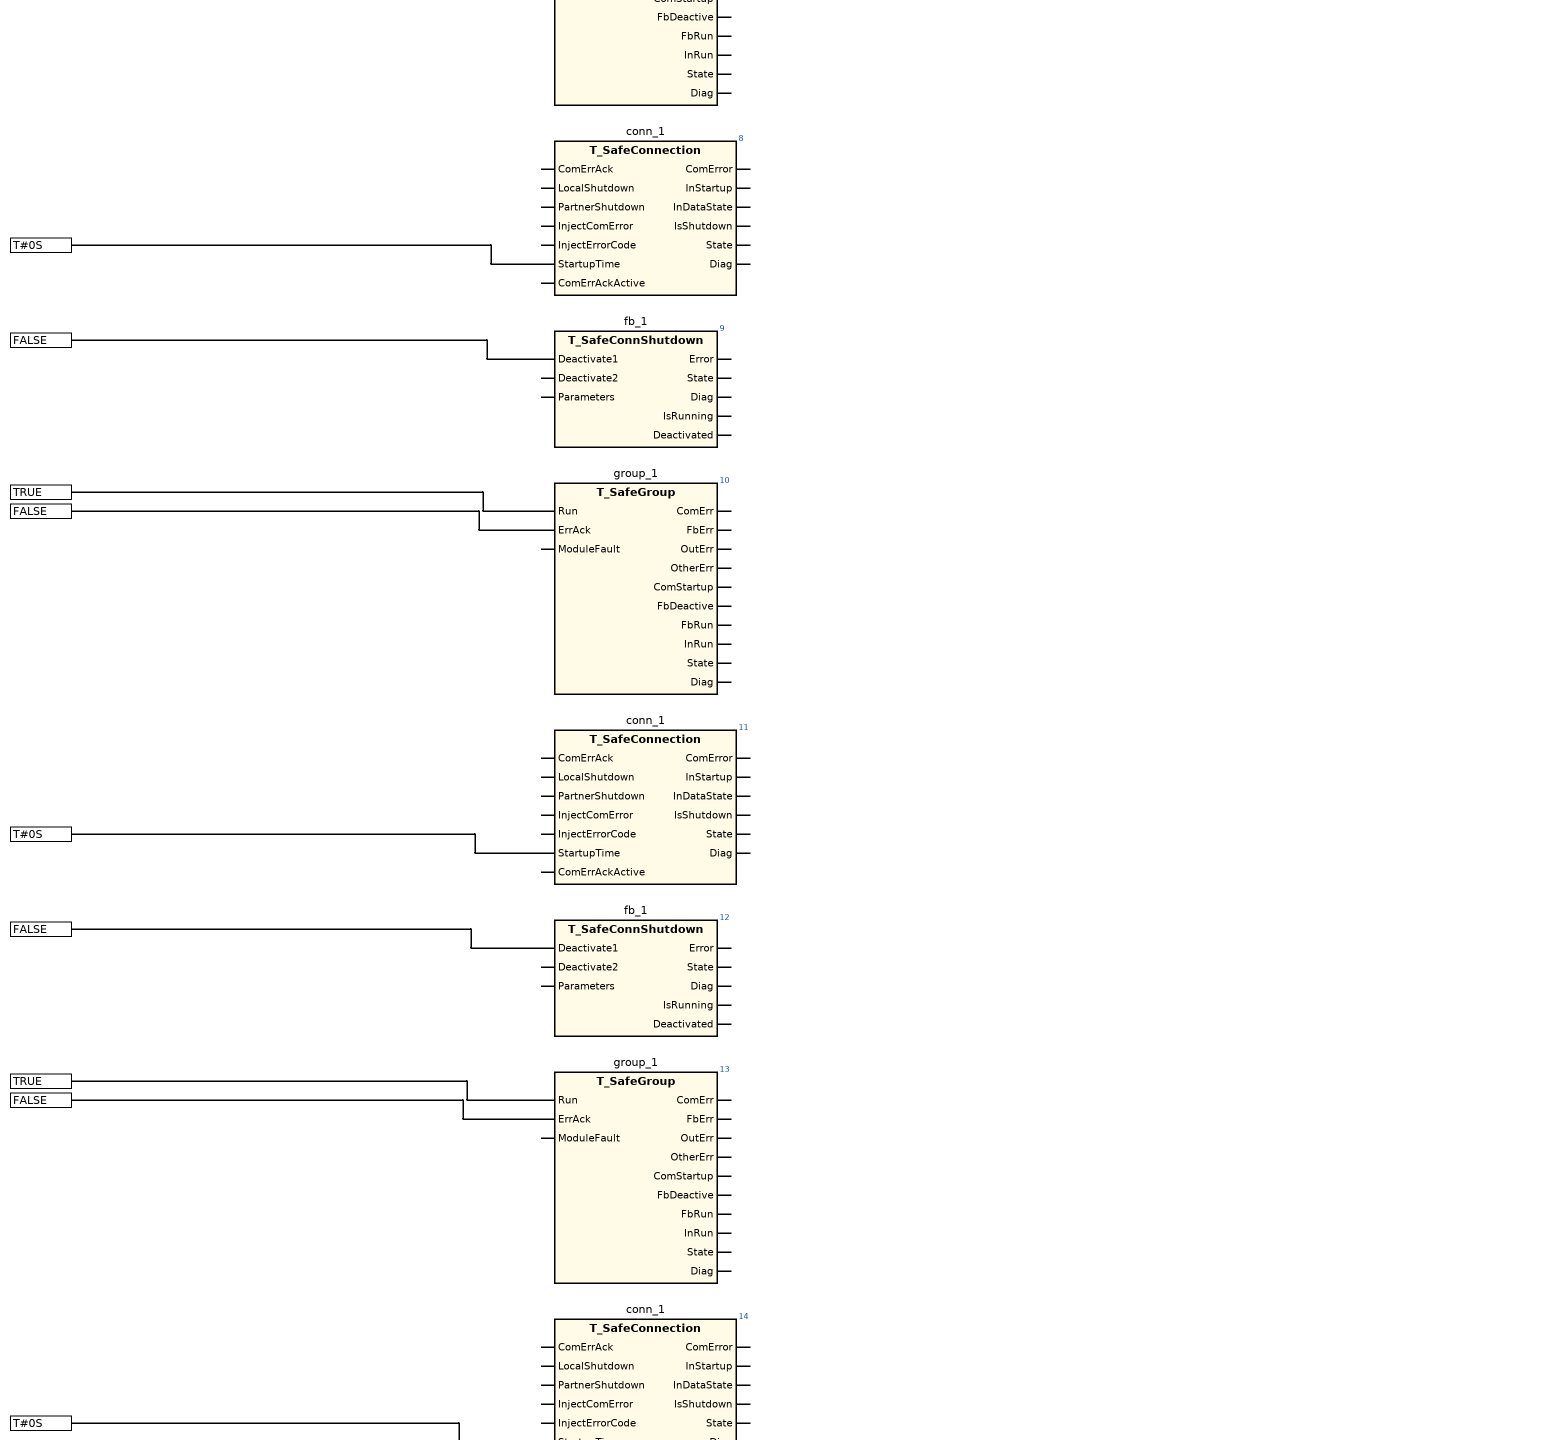
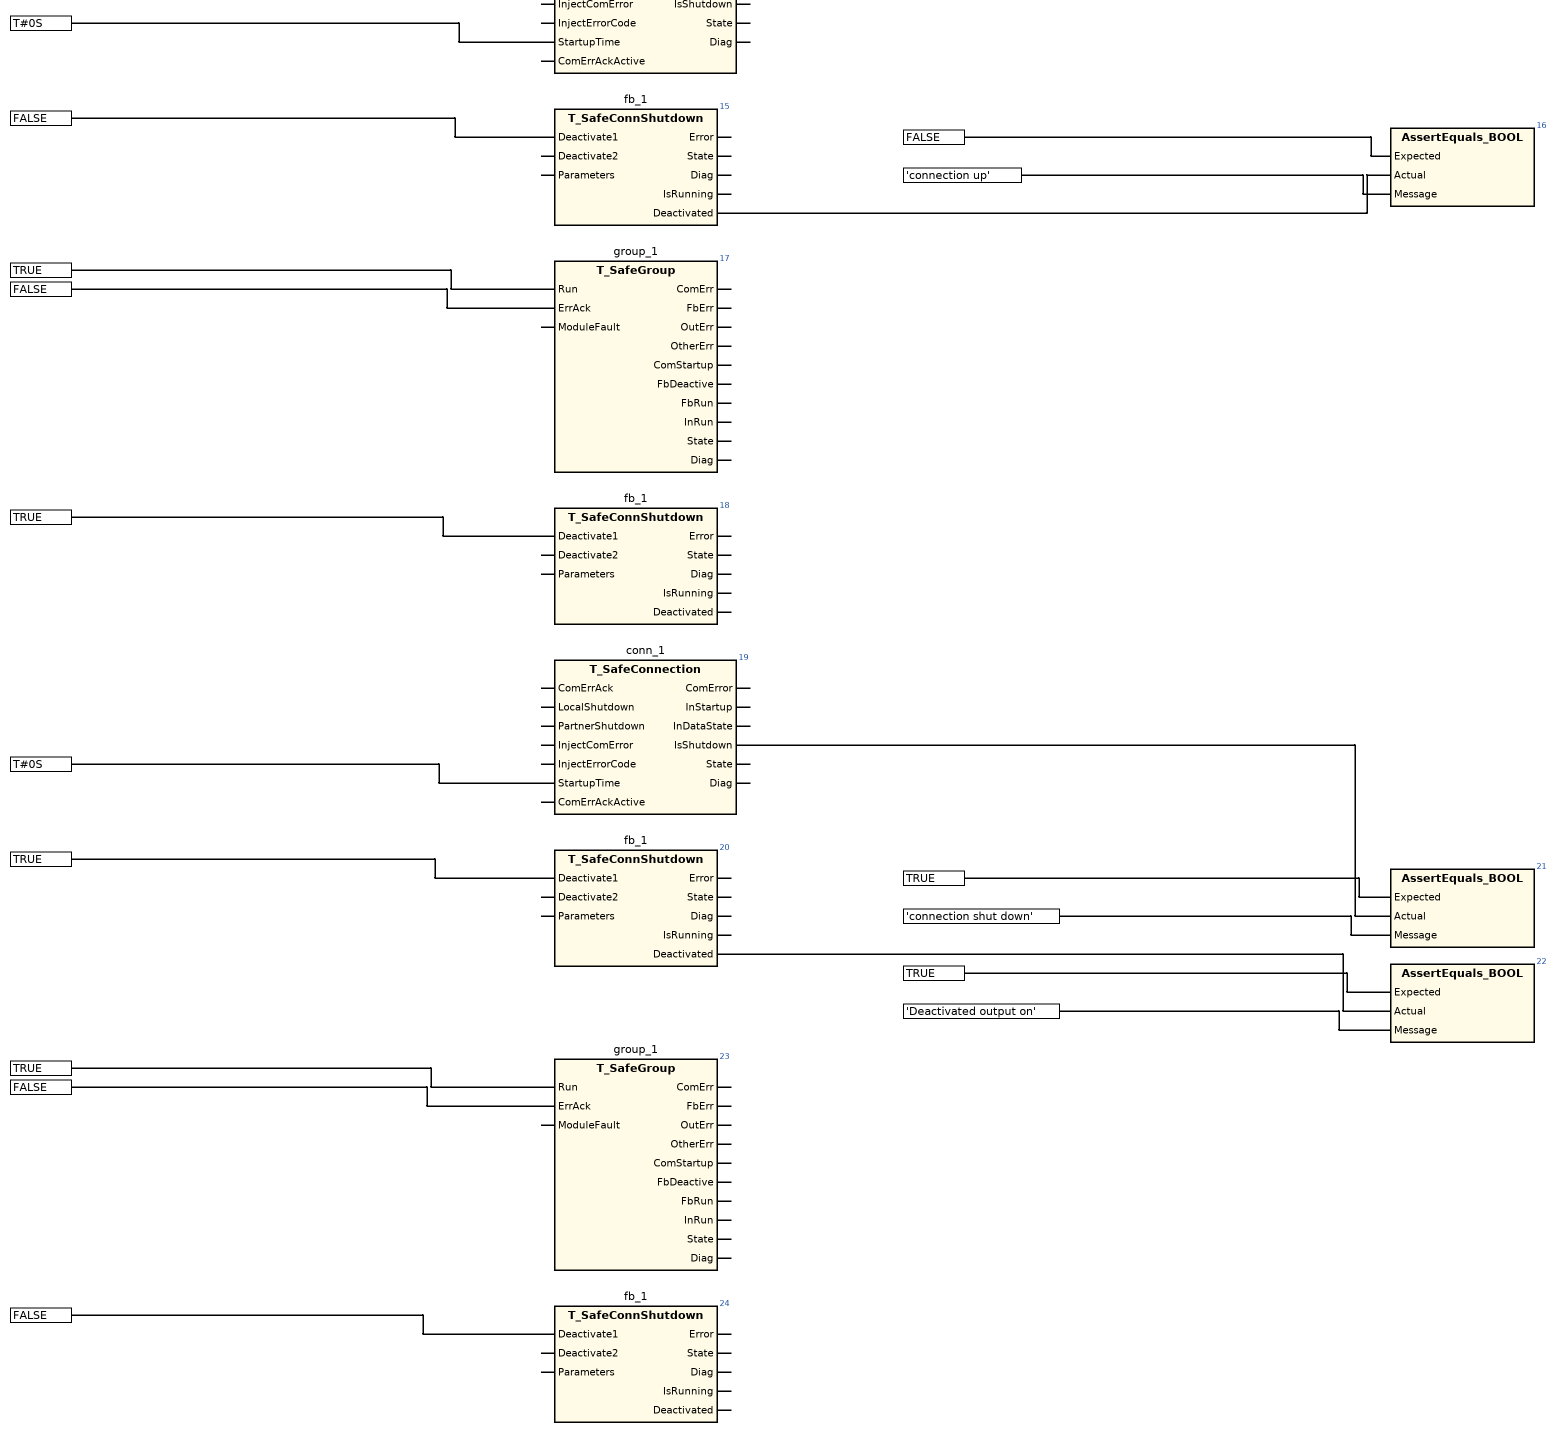
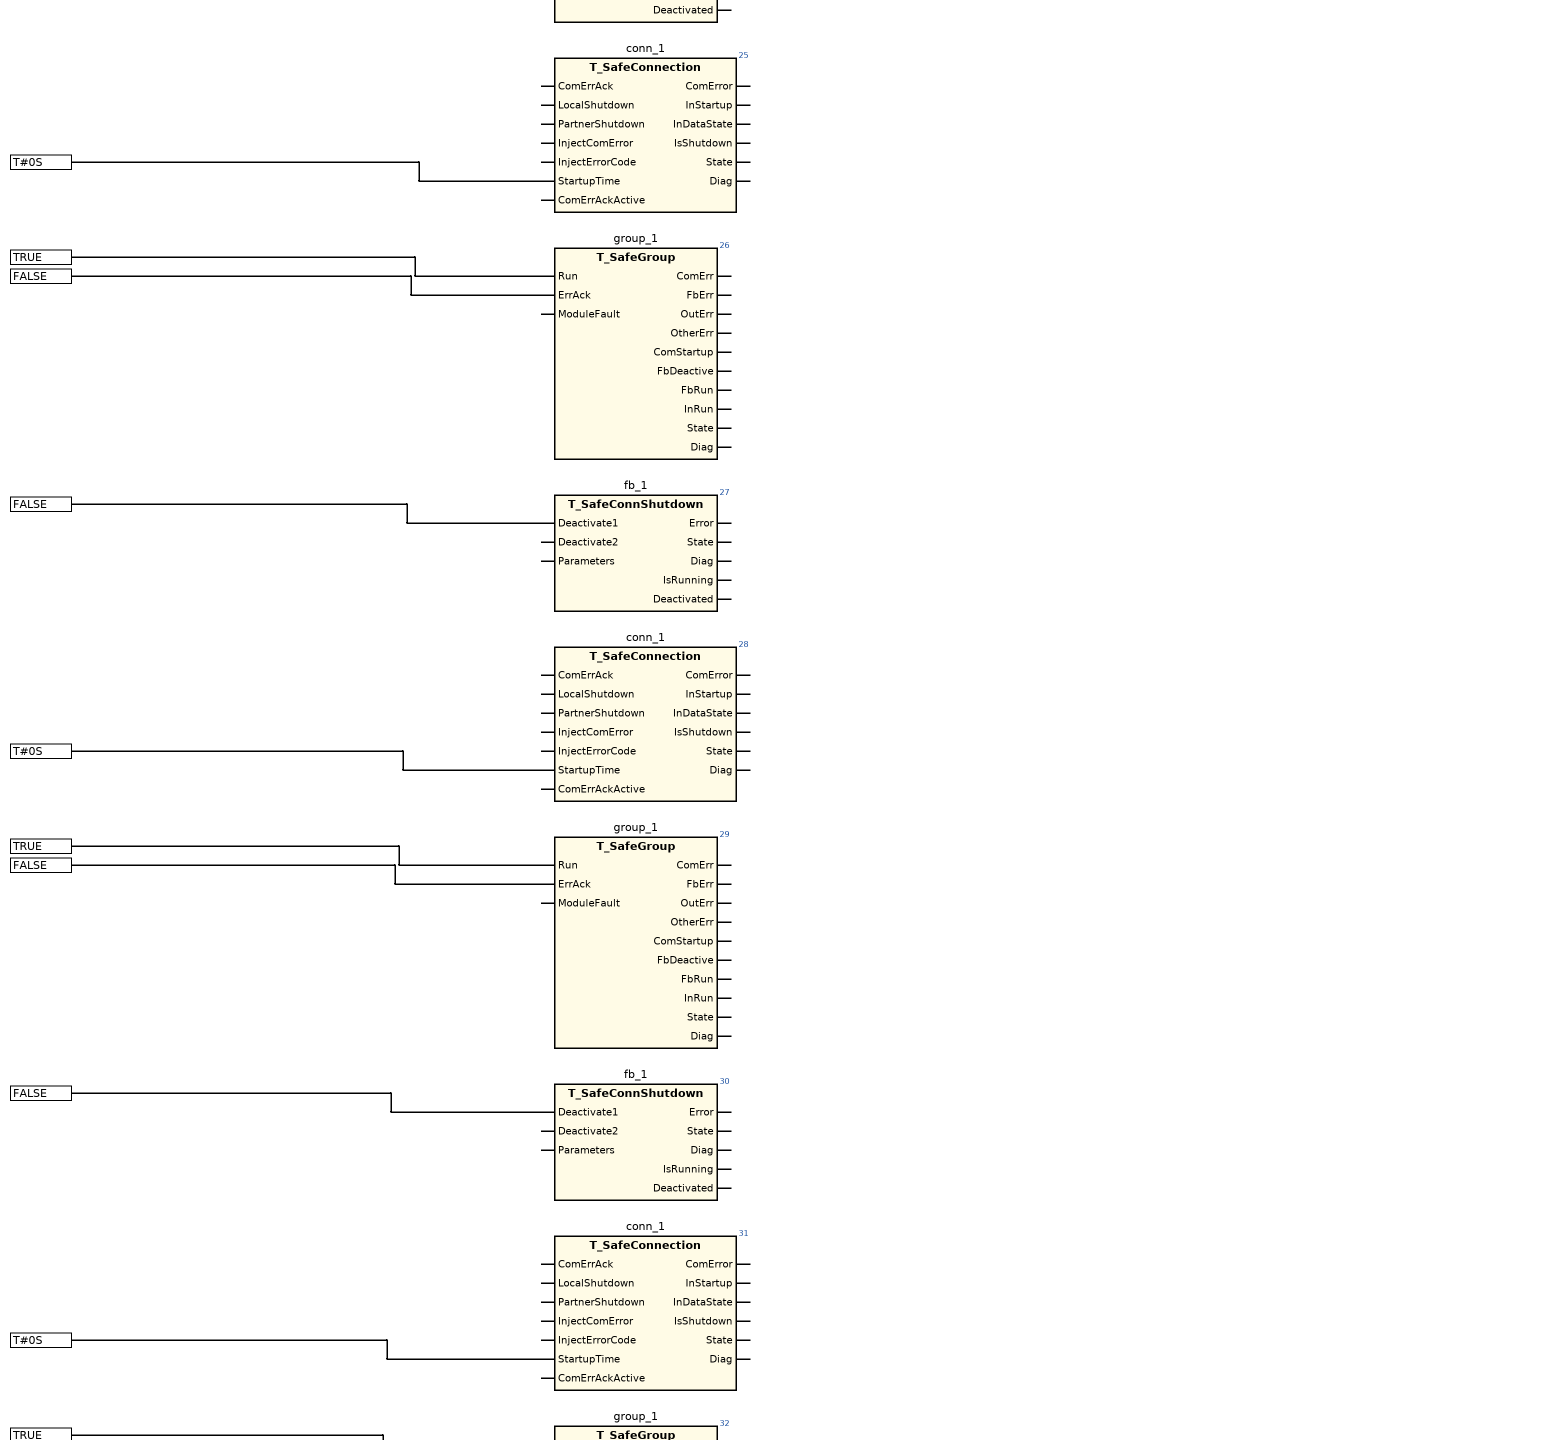
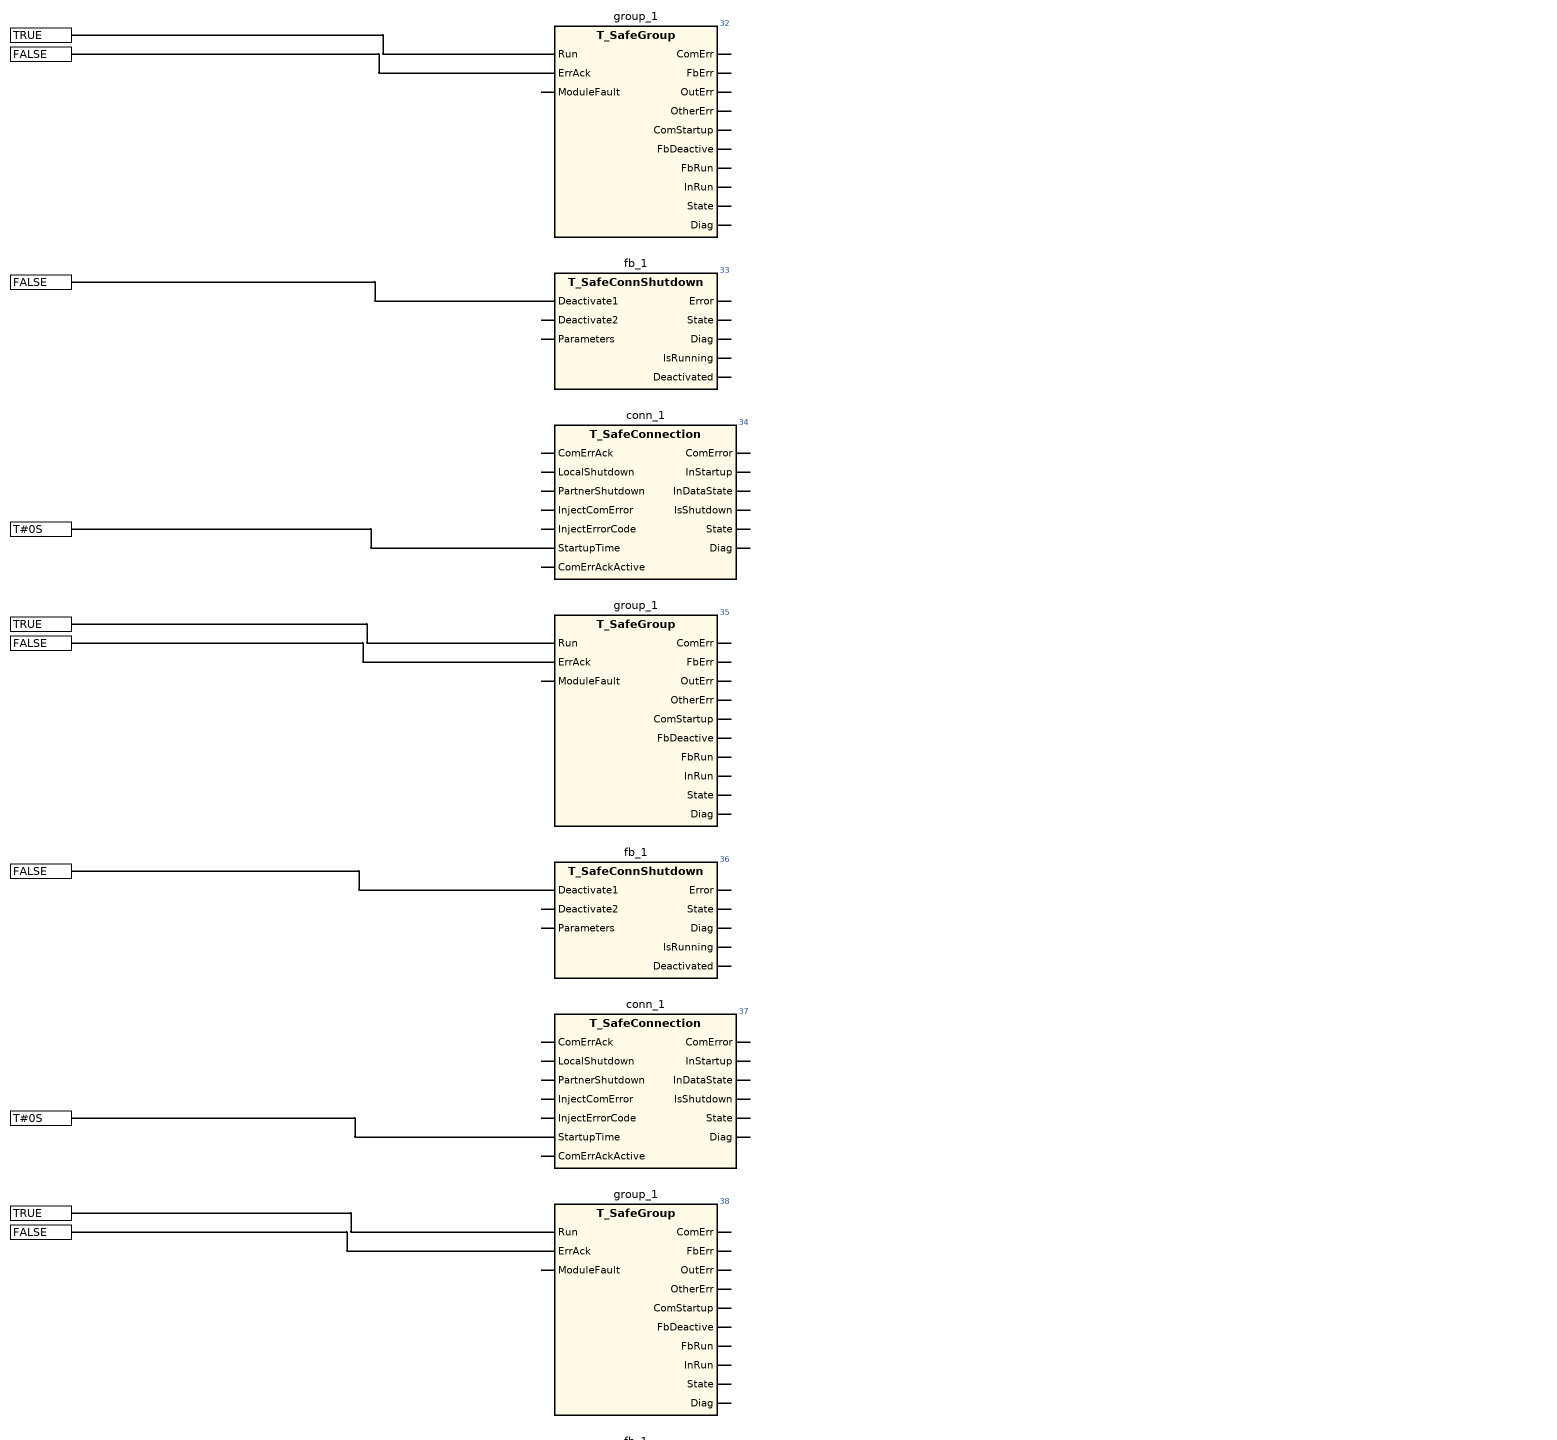
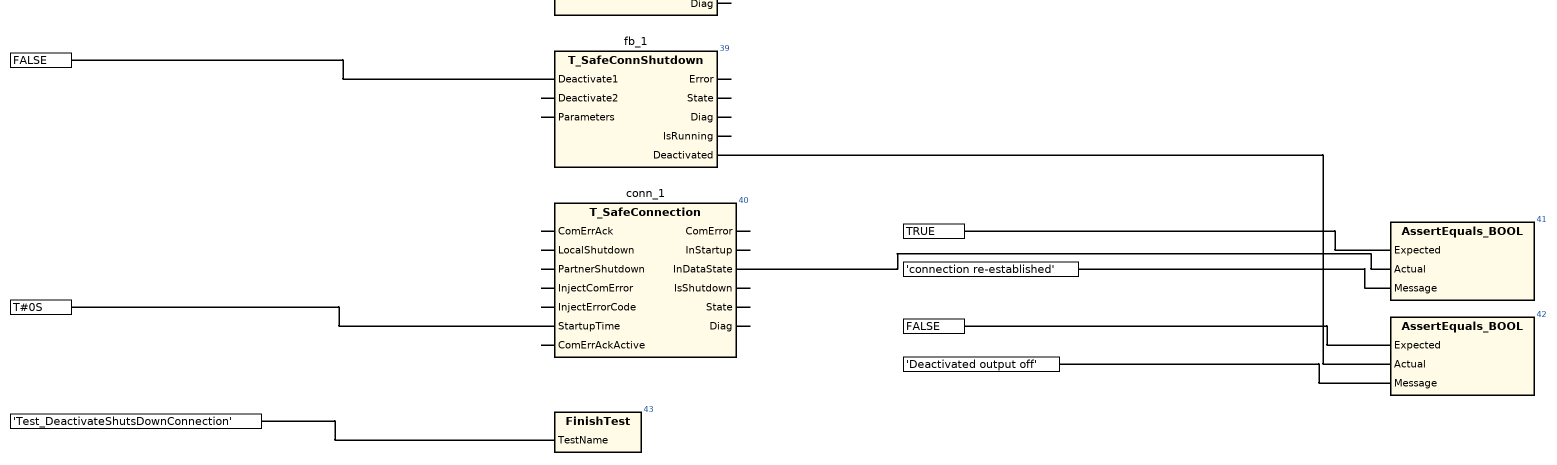
StartTest(TestName := 'Test_DeactivateShutsDownConnection');
group_1(Run := TRUE, ErrAck := FALSE); // T_SafeGroup
conn_1(StartupTime := T#0S); // T_SafeConnection
fb_1(Deactivate1 := FALSE); // T_SafeConnShutdown
group_1(Run := TRUE, ErrAck := FALSE); // T_SafeGroup
conn_1(StartupTime := T#0S); // T_SafeConnection
fb_1(Deactivate1 := FALSE); // T_SafeConnShutdown
group_1(Run := TRUE, ErrAck := FALSE); // T_SafeGroup
conn_1(StartupTime := T#0S); // T_SafeConnection
fb_1(Deactivate1 := FALSE); // T_SafeConnShutdown
group_1(Run := TRUE, ErrAck := FALSE); // T_SafeGroup
conn_1(StartupTime := T#0S); // T_SafeConnection
fb_1(Deactivate1 := FALSE); // T_SafeConnShutdown
group_1(Run := TRUE, ErrAck := FALSE); // T_SafeGroup
conn_1(StartupTime := T#0S); // T_SafeConnection
fb_1(Deactivate1 := FALSE); // T_SafeConnShutdown
AssertEquals_BOOL(Expected := FALSE, Actual := fb_1.Deactivated, Message := 'connection up');
group_1(Run := TRUE, ErrAck := FALSE); // T_SafeGroup
fb_1(Deactivate1 := TRUE); // T_SafeConnShutdown
conn_1(StartupTime := T#0S); // T_SafeConnection
fb_1(Deactivate1 := TRUE); // T_SafeConnShutdown
AssertEquals_BOOL(Expected := TRUE, Actual := conn_1.IsShutdown, Message := 'connection shut down');
AssertEquals_BOOL(Expected := TRUE, Actual := fb_1.Deactivated, Message := 'Deactivated output on');
group_1(Run := TRUE, ErrAck := FALSE); // T_SafeGroup
fb_1(Deactivate1 := FALSE); // T_SafeConnShutdown
conn_1(StartupTime := T#0S); // T_SafeConnection
group_1(Run := TRUE, ErrAck := FALSE); // T_SafeGroup
fb_1(Deactivate1 := FALSE); // T_SafeConnShutdown
conn_1(StartupTime := T#0S); // T_SafeConnection
group_1(Run := TRUE, ErrAck := FALSE); // T_SafeGroup
fb_1(Deactivate1 := FALSE); // T_SafeConnShutdown
conn_1(StartupTime := T#0S); // T_SafeConnection
group_1(Run := TRUE, ErrAck := FALSE); // T_SafeGroup
fb_1(Deactivate1 := FALSE); // T_SafeConnShutdown
conn_1(StartupTime := T#0S); // T_SafeConnection
group_1(Run := TRUE, ErrAck := FALSE); // T_SafeGroup
fb_1(Deactivate1 := FALSE); // T_SafeConnShutdown
conn_1(StartupTime := T#0S); // T_SafeConnection
group_1(Run := TRUE, ErrAck := FALSE); // T_SafeGroup
fb_1(Deactivate1 := FALSE); // T_SafeConnShutdown
conn_1(StartupTime := T#0S); // T_SafeConnection
AssertEquals_BOOL(Expected := TRUE, Actual := conn_1.InDataState, Message := 'connection re-established');
AssertEquals_BOOL(Expected := FALSE, Actual := fb_1.Deactivated, Message := 'Deactivated output off');
FinishTest(TestName := 'Test_DeactivateShutsDownConnection');
END_METHOD

END_FUNCTION_BLOCK

// Tests/T_SafeGroup_Tests_CFC
    // CFC twin of T_SafeGroup_Tests: the same tests drawn as CFC diagrams, the way a TwinSAFE project is authored.
    FUNCTION_BLOCK T_SafeGroup_Tests_CFC EXTENDS T_SafeCfcTestSuite
    VAR
    // Test_StopWhenRunFalse
    group_1 : T_SafeGroup;
    fb_1 : T_SafeAnd(group := group_1);
    // Test_RunsFunctionBlocksWithoutConnections
    group_2 : T_SafeGroup;
    fb_2 : T_SafeAnd(group := group_2);
    // Test_FbErrorStopsGroupAndErrAckRecovers
    group_3 : T_SafeGroup;
    eStop_3 : T_SafeEStop(group := group_3);
    andFb_3 : T_SafeAnd(group := group_3);
    // Test_ConnectionStartupAndComError
    group_4 : T_SafeGroup;
    terminal_4 : T_SafeInputTerminal(group := group_4);
    t1a_4 : TON;
    t1b_4 : TON;
    t2b_4 : TON;
    trig1a_4 : R_TRIG;
    trig1b_4 : R_TRIG;
    trig2b_4 : R_TRIG;
    t3_4 : TON;
    trig3_4 : R_TRIG;
    t0_4 : TON;
    t1_4 : TON;
    t2_4 : TON;
    t4_4 : TON;
    trig0_4 : R_TRIG;
    trig1_4 : R_TRIG;
    trig2_4 : R_TRIG;
    trig4_4 : R_TRIG;
END_VAR

Test_StopWhenRunFalse();
Test_RunsFunctionBlocksWithoutConnections();
Test_FbErrorStopsGroupAndErrAckRecovers();
Test_ConnectionStartupAndComError();

METHOD PRIVATE Test_ConnectionStartupAndComError
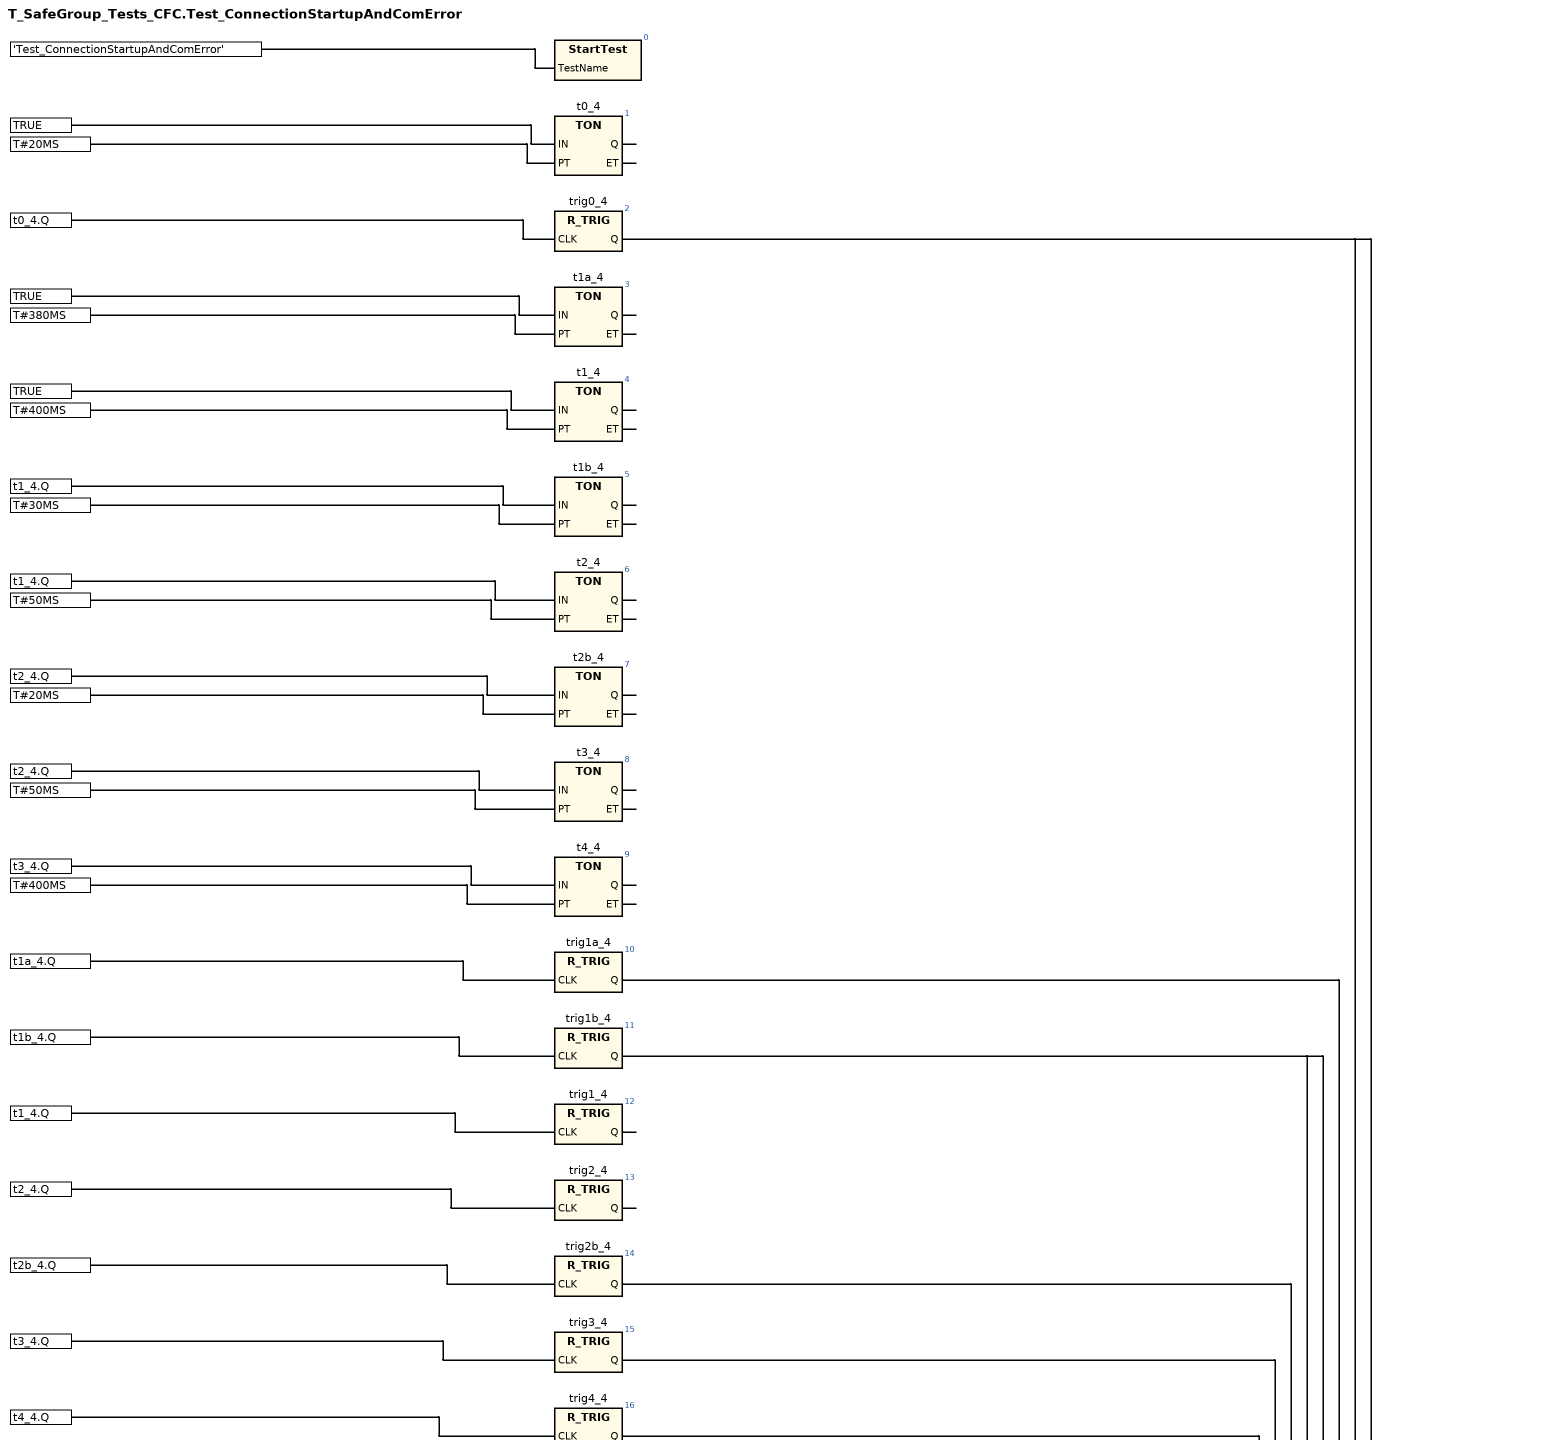
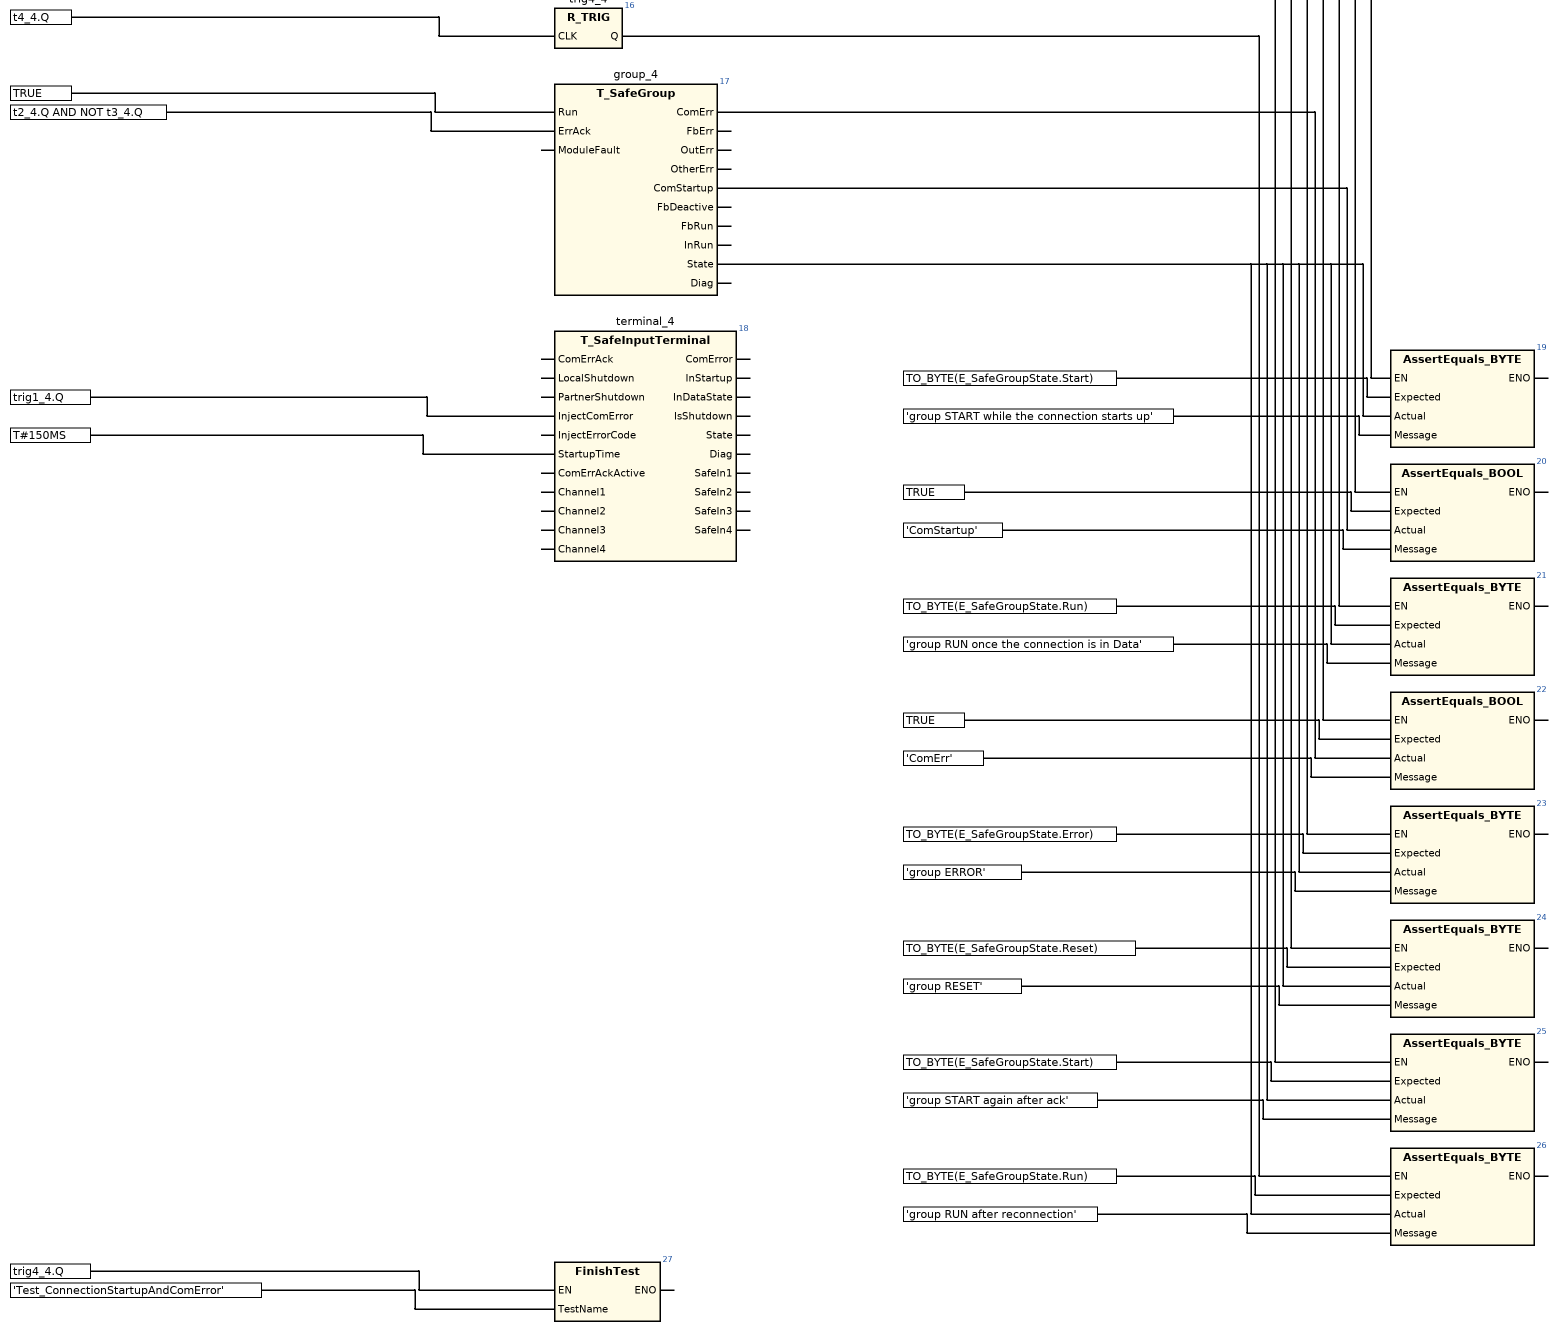
StartTest(TestName := 'Test_ConnectionStartupAndComError');
t0_4(IN := TRUE, PT := T#20MS); // TON
trig0_4(CLK := t0_4.Q); // R_TRIG
t1a_4(IN := TRUE, PT := T#380MS); // TON
t1_4(IN := TRUE, PT := T#400MS); // TON
t1b_4(IN := t1_4.Q, PT := T#30MS); // TON
t2_4(IN := t1_4.Q, PT := T#50MS); // TON
t2b_4(IN := t2_4.Q, PT := T#20MS); // TON
t3_4(IN := t2_4.Q, PT := T#50MS); // TON
t4_4(IN := t3_4.Q, PT := T#400MS); // TON
trig1a_4(CLK := t1a_4.Q); // R_TRIG
trig1b_4(CLK := t1b_4.Q); // R_TRIG
trig1_4(CLK := t1_4.Q); // R_TRIG
trig2_4(CLK := t2_4.Q); // R_TRIG
trig2b_4(CLK := t2b_4.Q); // R_TRIG
trig3_4(CLK := t3_4.Q); // R_TRIG
trig4_4(CLK := t4_4.Q); // R_TRIG
group_4(Run := TRUE, ErrAck := t2_4.Q AND NOT t3_4.Q); // T_SafeGroup
terminal_4(InjectComError := trig1_4.Q, StartupTime := T#150MS); // T_SafeInputTerminal
IF trig0_4.Q THEN AssertEquals_BYTE(Expected := TO_BYTE(E_SafeGroupState.Start), Actual := group_4.State, Message := 'group START while the connection starts up'); END_IF
IF trig0_4.Q THEN AssertEquals_BOOL(Expected := TRUE, Actual := group_4.ComStartup, Message := 'ComStartup'); END_IF
IF trig1a_4.Q THEN AssertEquals_BYTE(Expected := TO_BYTE(E_SafeGroupState.Run), Actual := group_4.State, Message := 'group RUN once the connection is in Data'); END_IF
IF trig1b_4.Q THEN AssertEquals_BOOL(Expected := TRUE, Actual := group_4.ComErr, Message := 'ComErr'); END_IF
IF trig1b_4.Q THEN AssertEquals_BYTE(Expected := TO_BYTE(E_SafeGroupState.Error), Actual := group_4.State, Message := 'group ERROR'); END_IF
IF trig2b_4.Q THEN AssertEquals_BYTE(Expected := TO_BYTE(E_SafeGroupState.Reset), Actual := group_4.State, Message := 'group RESET'); END_IF
IF trig3_4.Q THEN AssertEquals_BYTE(Expected := TO_BYTE(E_SafeGroupState.Start), Actual := group_4.State, Message := 'group START again after ack'); END_IF
IF trig4_4.Q THEN AssertEquals_BYTE(Expected := TO_BYTE(E_SafeGroupState.Run), Actual := group_4.State, Message := 'group RUN after reconnection'); END_IF
IF trig4_4.Q THEN FinishTest(TestName := 'Test_ConnectionStartupAndComError'); END_IF
END_METHOD

METHOD PRIVATE Test_FbErrorStopsGroupAndErrAckRecovers
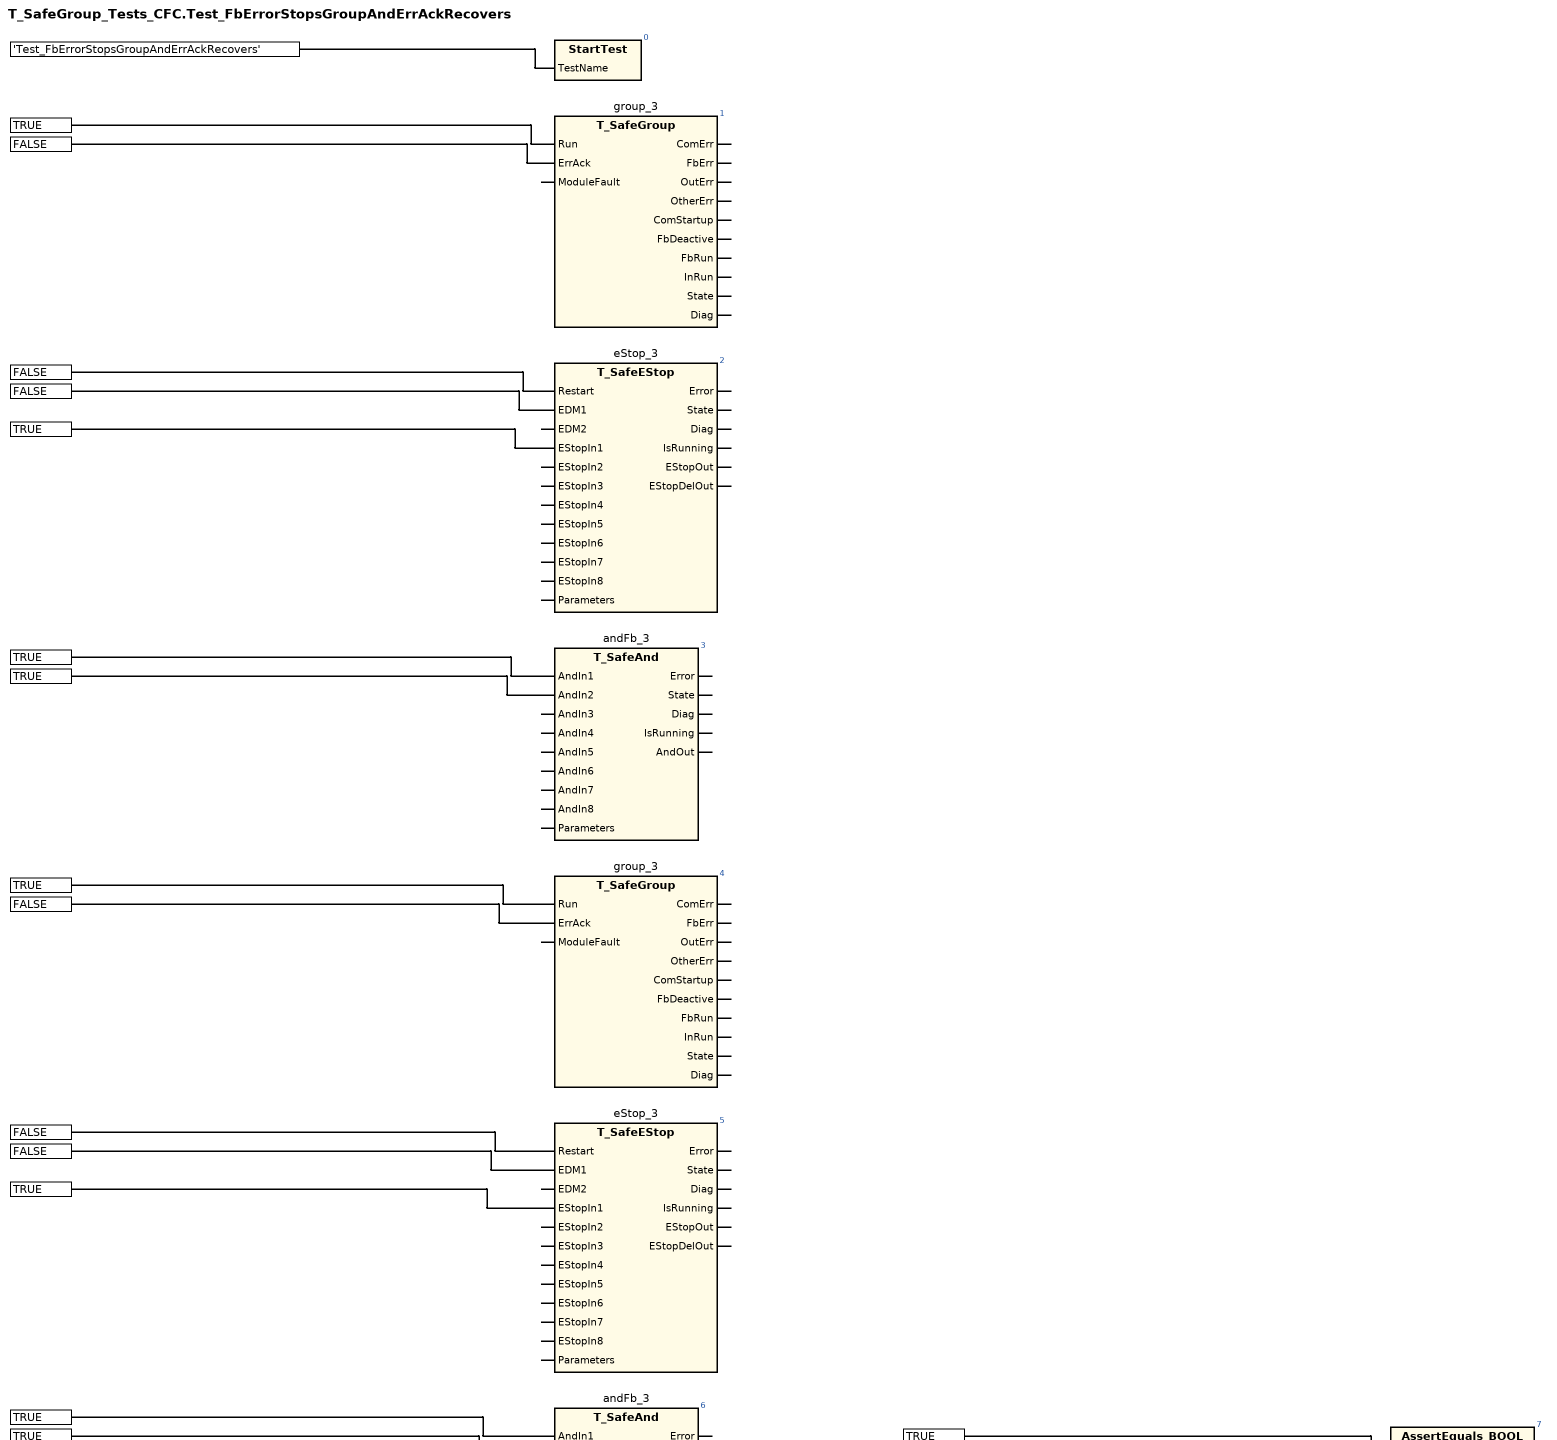
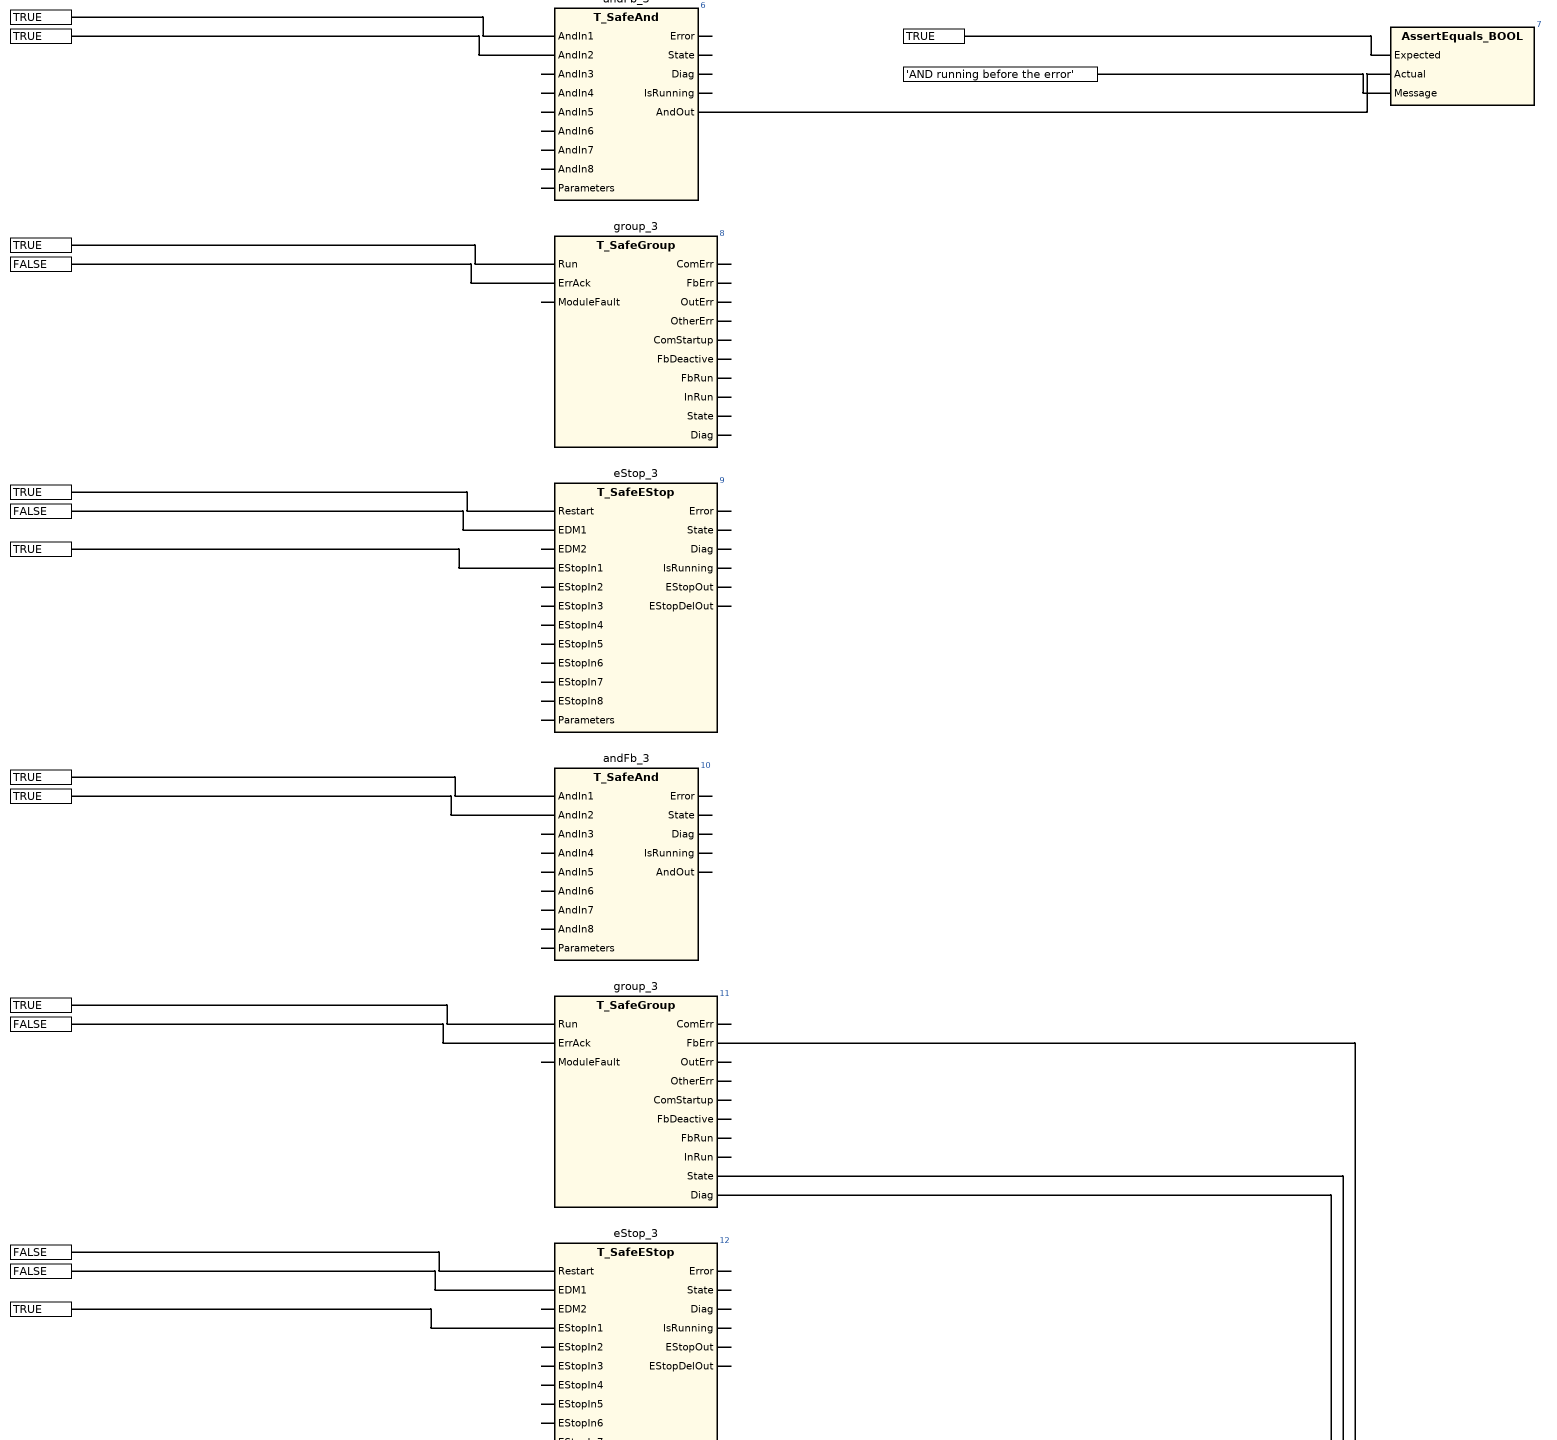
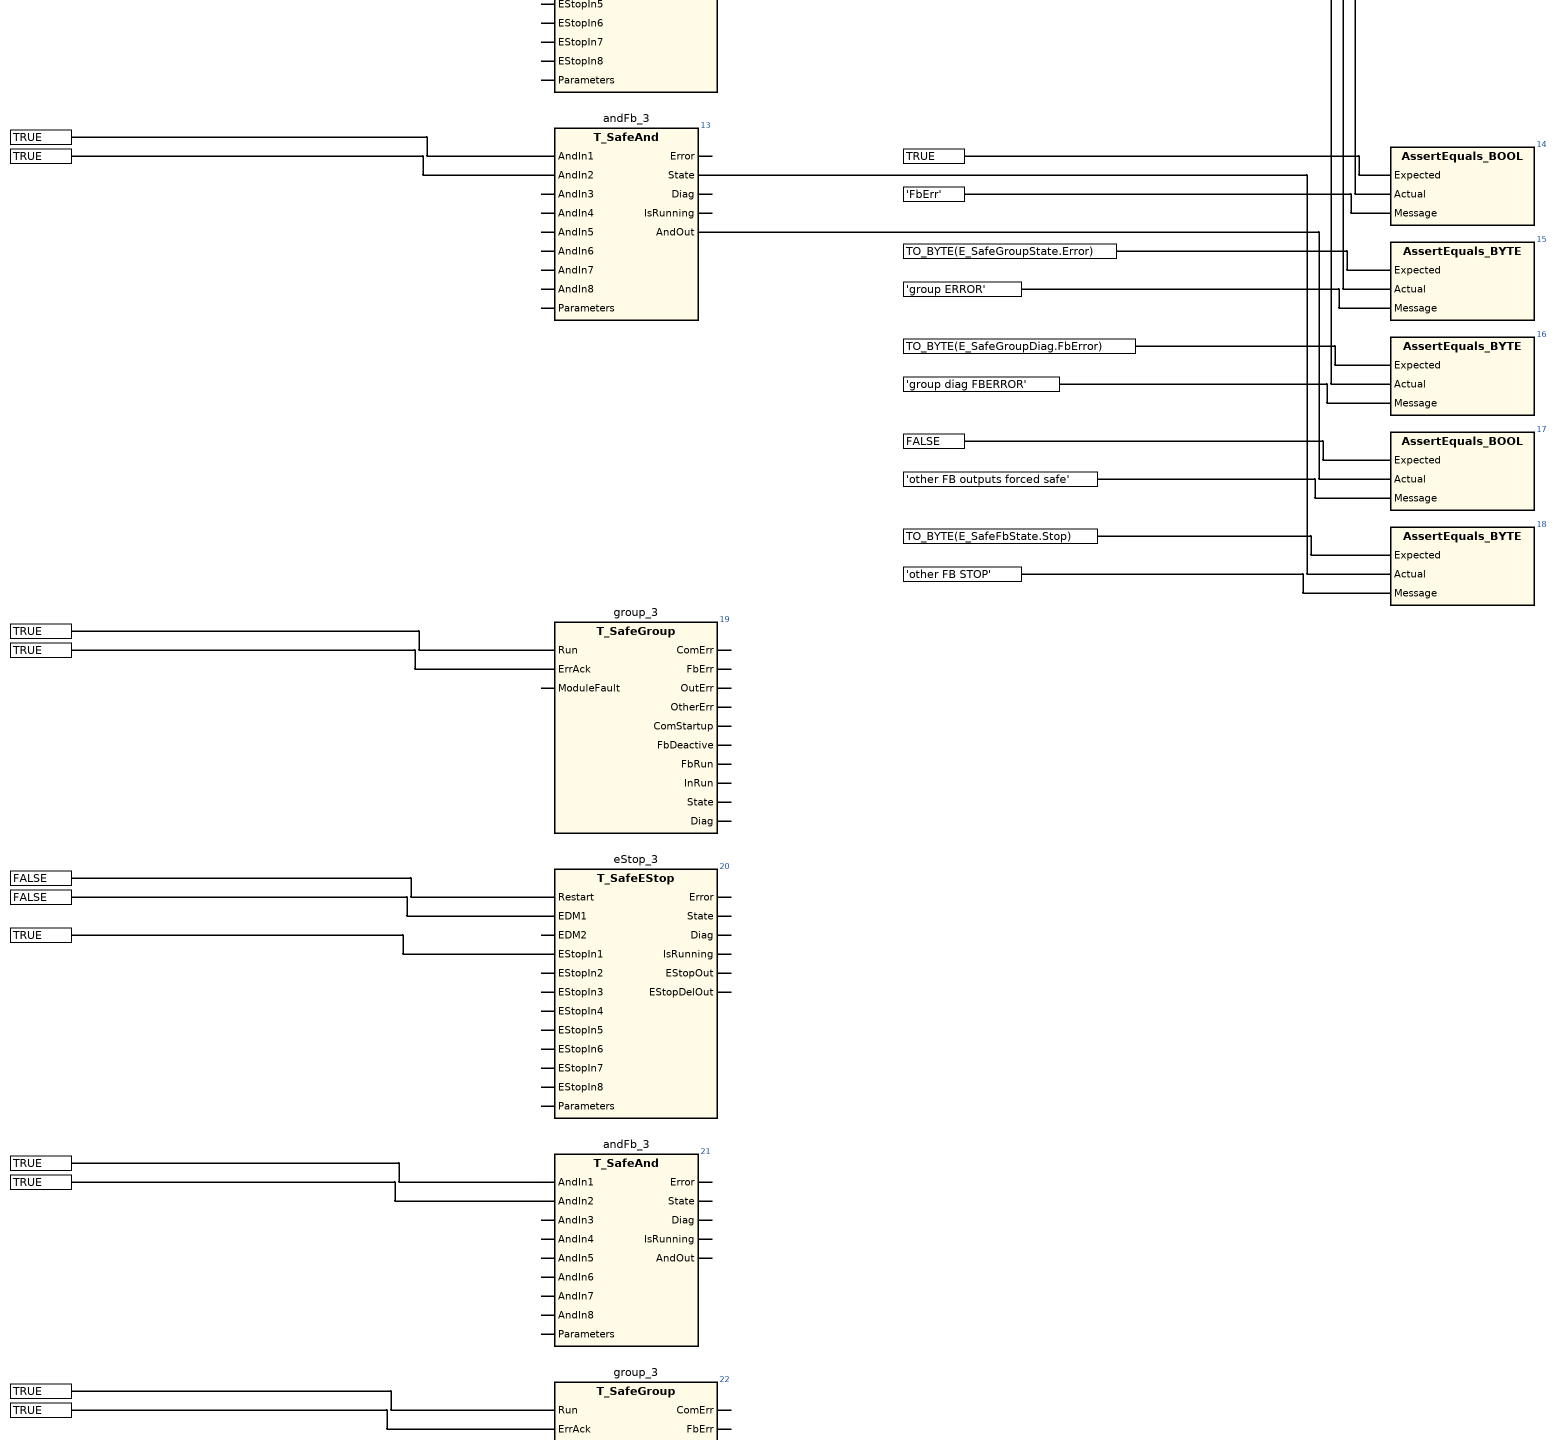
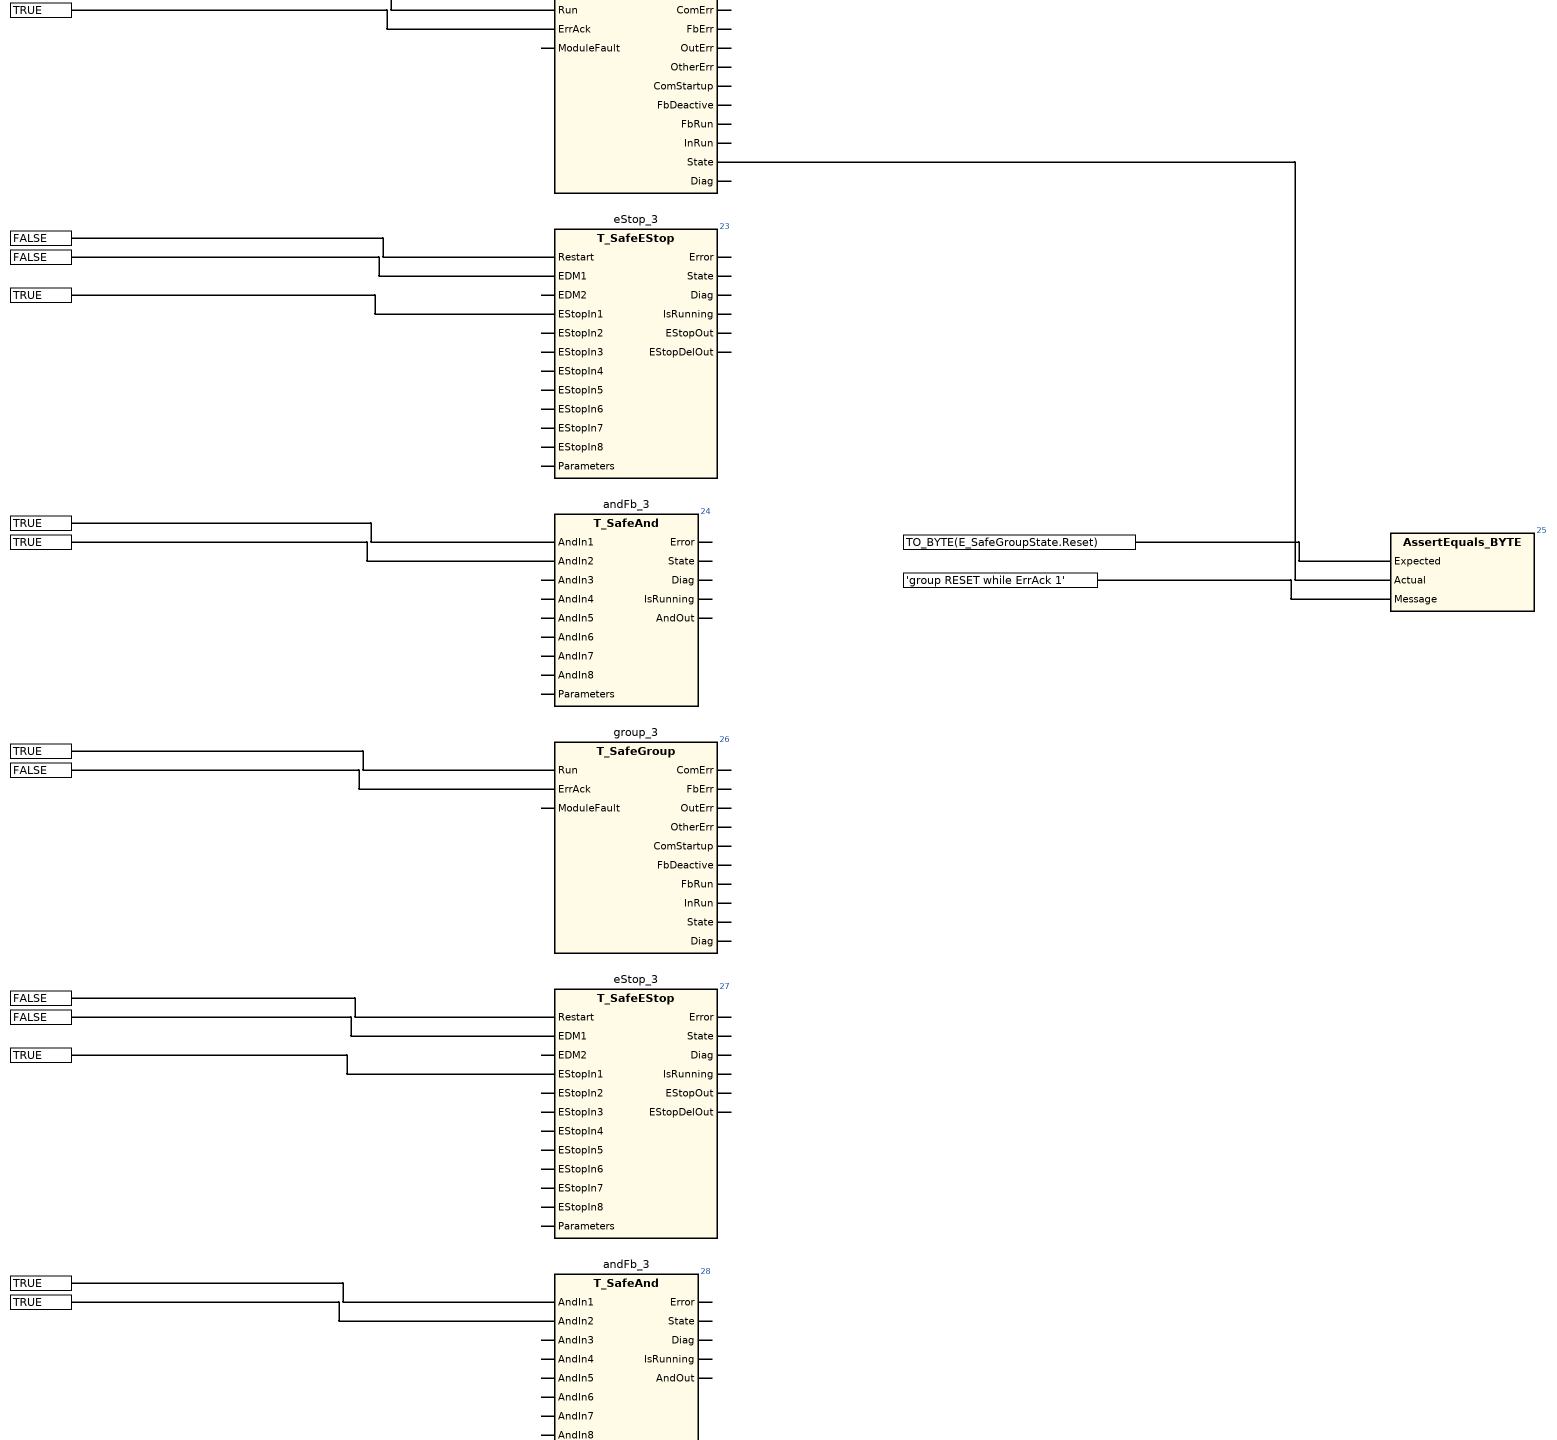
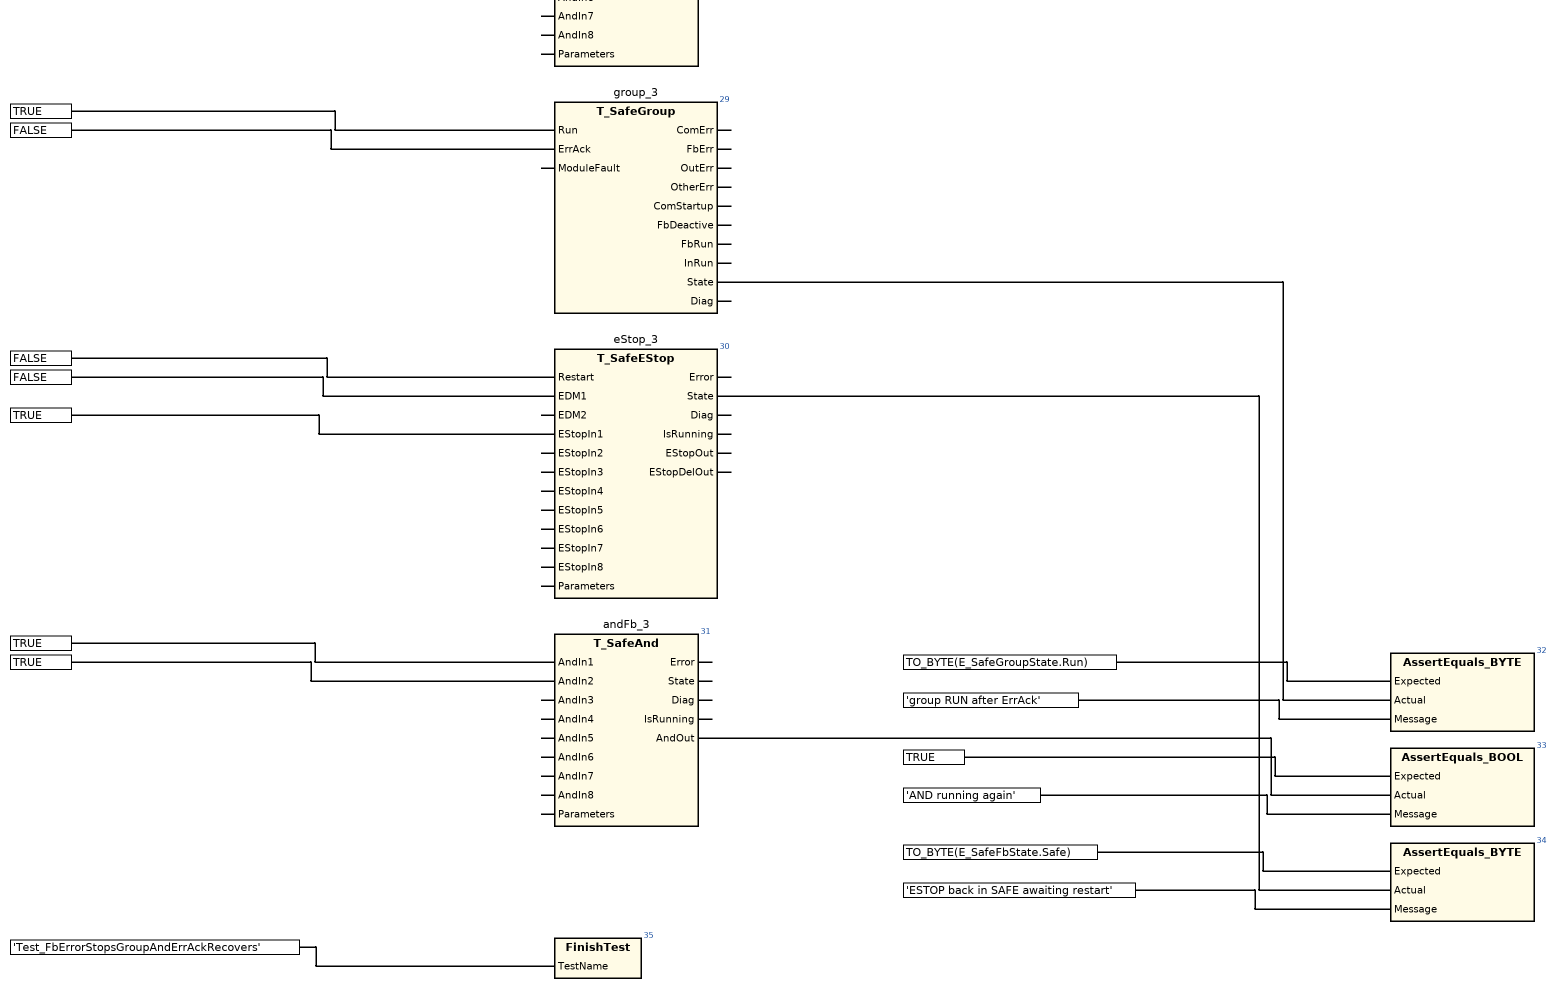
StartTest(TestName := 'Test_FbErrorStopsGroupAndErrAckRecovers');
group_3(Run := TRUE, ErrAck := FALSE); // T_SafeGroup
eStop_3(Restart := FALSE, EDM1 := FALSE, EStopIn1 := TRUE); // T_SafeEStop
andFb_3(AndIn1 := TRUE, AndIn2 := TRUE); // T_SafeAnd
group_3(Run := TRUE, ErrAck := FALSE); // T_SafeGroup
eStop_3(Restart := FALSE, EDM1 := FALSE, EStopIn1 := TRUE); // T_SafeEStop
andFb_3(AndIn1 := TRUE, AndIn2 := TRUE); // T_SafeAnd
AssertEquals_BOOL(Expected := TRUE, Actual := andFb_3.AndOut, Message := 'AND running before the error');
group_3(Run := TRUE, ErrAck := FALSE); // T_SafeGroup
eStop_3(Restart := TRUE, EDM1 := FALSE, EStopIn1 := TRUE); // T_SafeEStop
andFb_3(AndIn1 := TRUE, AndIn2 := TRUE); // T_SafeAnd
group_3(Run := TRUE, ErrAck := FALSE); // T_SafeGroup
eStop_3(Restart := FALSE, EDM1 := FALSE, EStopIn1 := TRUE); // T_SafeEStop
andFb_3(AndIn1 := TRUE, AndIn2 := TRUE); // T_SafeAnd
AssertEquals_BOOL(Expected := TRUE, Actual := group_3.FbErr, Message := 'FbErr');
AssertEquals_BYTE(Expected := TO_BYTE(E_SafeGroupState.Error), Actual := group_3.State, Message := 'group ERROR');
AssertEquals_BYTE(Expected := TO_BYTE(E_SafeGroupDiag.FbError), Actual := group_3.Diag, Message := 'group diag FBERROR');
AssertEquals_BOOL(Expected := FALSE, Actual := andFb_3.AndOut, Message := 'other FB outputs forced safe');
AssertEquals_BYTE(Expected := TO_BYTE(E_SafeFbState.Stop), Actual := andFb_3.State, Message := 'other FB STOP');
group_3(Run := TRUE, ErrAck := TRUE); // T_SafeGroup
eStop_3(Restart := FALSE, EDM1 := FALSE, EStopIn1 := TRUE); // T_SafeEStop
andFb_3(AndIn1 := TRUE, AndIn2 := TRUE); // T_SafeAnd
group_3(Run := TRUE, ErrAck := TRUE); // T_SafeGroup
eStop_3(Restart := FALSE, EDM1 := FALSE, EStopIn1 := TRUE); // T_SafeEStop
andFb_3(AndIn1 := TRUE, AndIn2 := TRUE); // T_SafeAnd
AssertEquals_BYTE(Expected := TO_BYTE(E_SafeGroupState.Reset), Actual := group_3.State, Message := 'group RESET while ErrAck 1');
group_3(Run := TRUE, ErrAck := FALSE); // T_SafeGroup
eStop_3(Restart := FALSE, EDM1 := FALSE, EStopIn1 := TRUE); // T_SafeEStop
andFb_3(AndIn1 := TRUE, AndIn2 := TRUE); // T_SafeAnd
group_3(Run := TRUE, ErrAck := FALSE); // T_SafeGroup
eStop_3(Restart := FALSE, EDM1 := FALSE, EStopIn1 := TRUE); // T_SafeEStop
andFb_3(AndIn1 := TRUE, AndIn2 := TRUE); // T_SafeAnd
AssertEquals_BYTE(Expected := TO_BYTE(E_SafeGroupState.Run), Actual := group_3.State, Message := 'group RUN after ErrAck');
AssertEquals_BOOL(Expected := TRUE, Actual := andFb_3.AndOut, Message := 'AND running again');
AssertEquals_BYTE(Expected := TO_BYTE(E_SafeFbState.Safe), Actual := eStop_3.State, Message := 'ESTOP back in SAFE awaiting restart');
FinishTest(TestName := 'Test_FbErrorStopsGroupAndErrAckRecovers');
END_METHOD

METHOD PRIVATE Test_RunsFunctionBlocksWithoutConnections
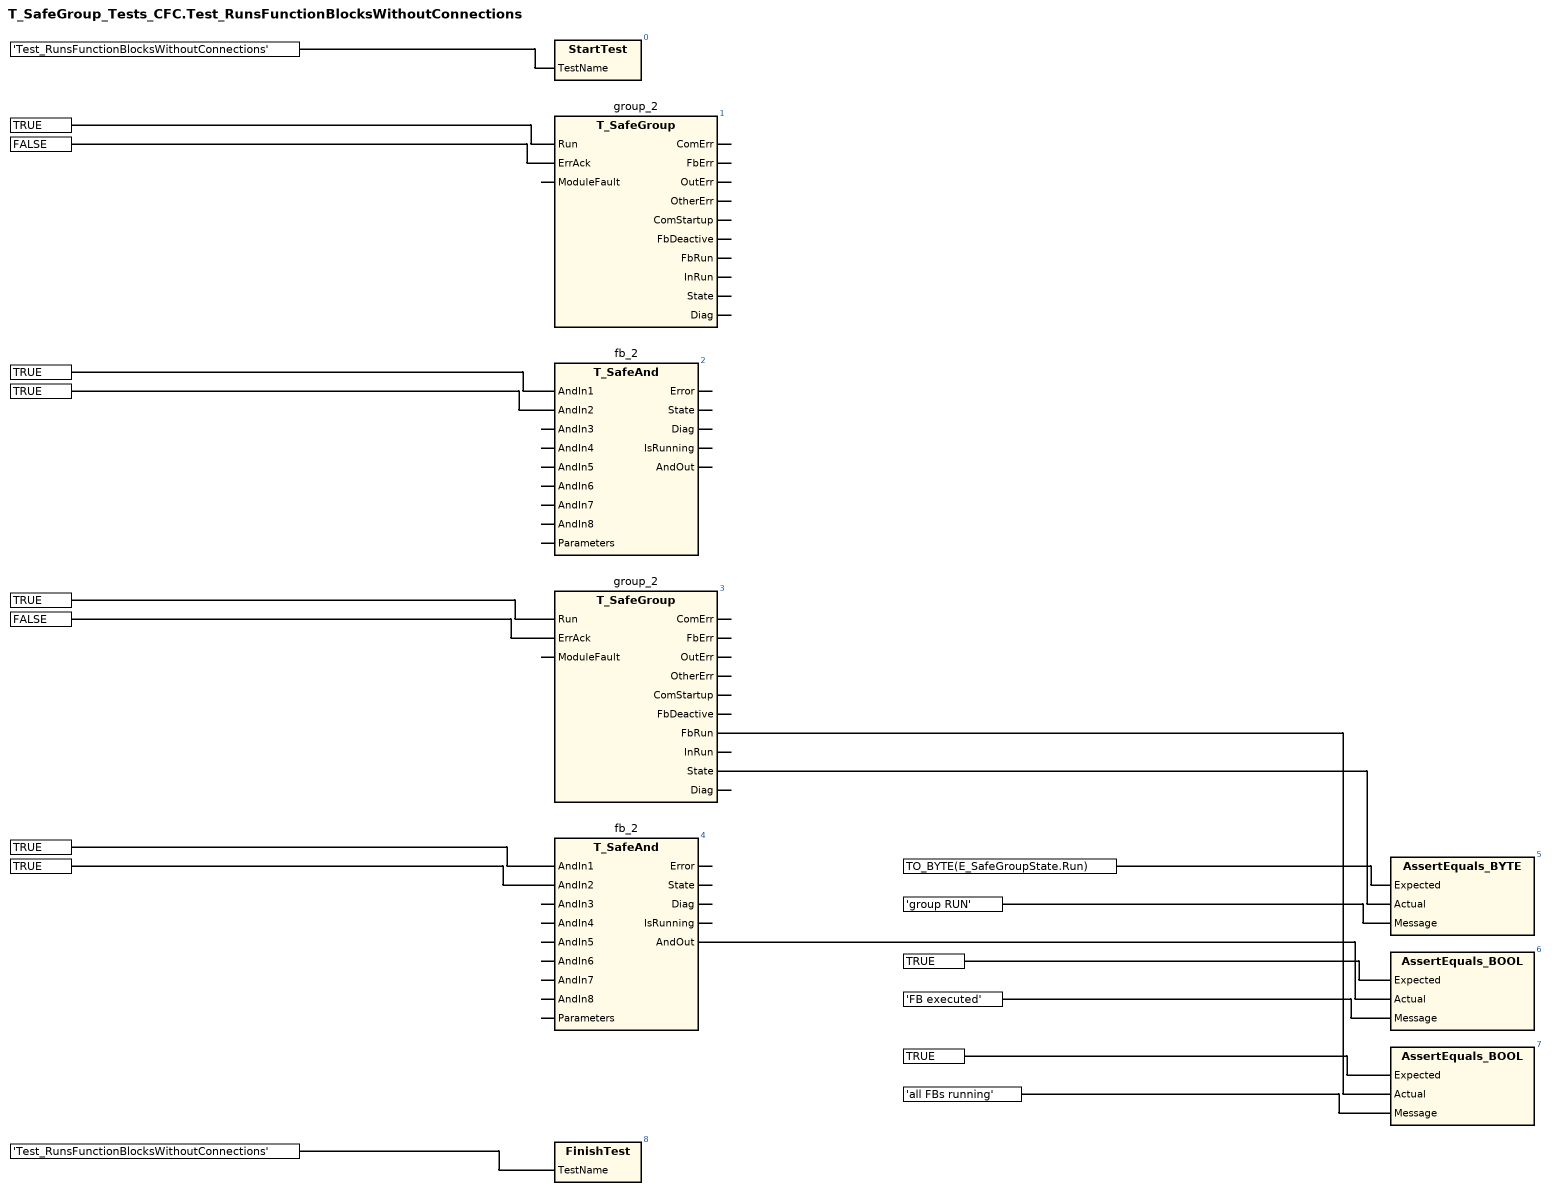
StartTest(TestName := 'Test_RunsFunctionBlocksWithoutConnections');
group_2(Run := TRUE, ErrAck := FALSE); // T_SafeGroup
fb_2(AndIn1 := TRUE, AndIn2 := TRUE); // T_SafeAnd
group_2(Run := TRUE, ErrAck := FALSE); // T_SafeGroup
fb_2(AndIn1 := TRUE, AndIn2 := TRUE); // T_SafeAnd
AssertEquals_BYTE(Expected := TO_BYTE(E_SafeGroupState.Run), Actual := group_2.State, Message := 'group RUN');
AssertEquals_BOOL(Expected := TRUE, Actual := fb_2.AndOut, Message := 'FB executed');
AssertEquals_BOOL(Expected := TRUE, Actual := group_2.FbRun, Message := 'all FBs running');
FinishTest(TestName := 'Test_RunsFunctionBlocksWithoutConnections');
END_METHOD

METHOD PRIVATE Test_StopWhenRunFalse
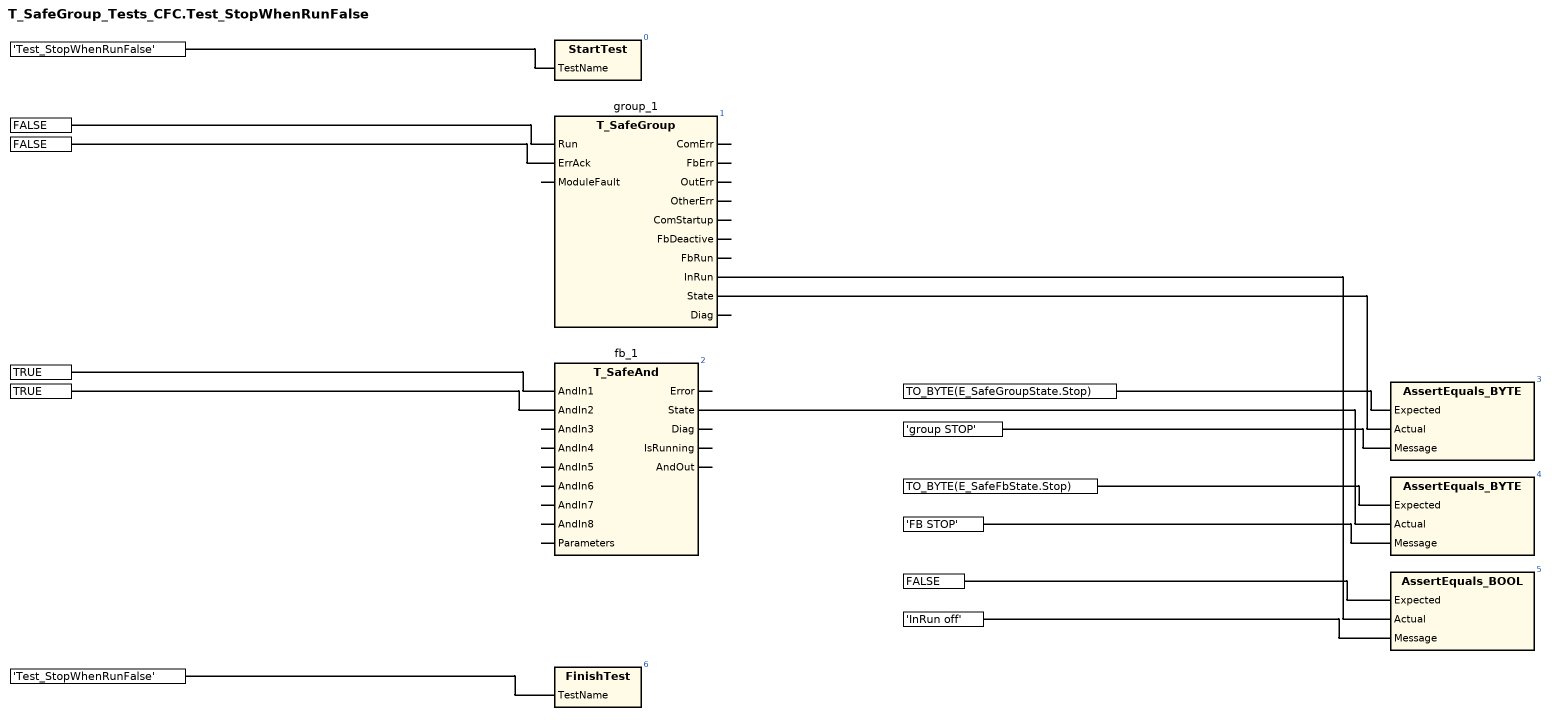
StartTest(TestName := 'Test_StopWhenRunFalse');
group_1(Run := FALSE, ErrAck := FALSE); // T_SafeGroup
fb_1(AndIn1 := TRUE, AndIn2 := TRUE); // T_SafeAnd
AssertEquals_BYTE(Expected := TO_BYTE(E_SafeGroupState.Stop), Actual := group_1.State, Message := 'group STOP');
AssertEquals_BYTE(Expected := TO_BYTE(E_SafeFbState.Stop), Actual := fb_1.State, Message := 'FB STOP');
AssertEquals_BOOL(Expected := FALSE, Actual := group_1.InRun, Message := 'InRun off');
FinishTest(TestName := 'Test_StopWhenRunFalse');
END_METHOD

END_FUNCTION_BLOCK
